(* PLC project forms.project, CODESYS CODESYS V3.5 SP17 Patch 3 *)
(* stored: creationDateTime 2026-10-20T03:44:11.3044873, modificationDateTime 1601-01-01T03:00:00 *)

TYPE ST_Probe : STRUCT
  a : INT;
  b : BOOL;
END_STRUCT;
END_TYPE
